(* CODESYS project festo_cmmt_as_etc.library
   DefaultNamespace: KOSTAL.TC3.Device.Axis.FESTO.CMMT_AS.ETC
   DocFormat: reStructuredText
   Description: Library to handle the FESTO CMMT_AS axis controller via EtherCAT
   Author: A.Zajic
   Title: KOSTAL.TC3.Device.Axis.FESTO.CMMT_AS.ETC
   Version: 2019.0.0.0
   Company: KOSTAL GmbH & Co.KG
   Placeholder: KOSTAL.TC3.Device.Axis.FESTO.CMMT_AS.ETC

Project tree, tasks and I/O mapping:
  libraries: Festo_PtP_Base, 3.5.15.32 (Festo); Festo_PtP_CiA402, 3.5.15.32 (Festo); Festo_PtP_CiA402_ETC, 3.5.15.32 (Festo); Festo_PtP_CiA402_ETC_CMMT_AS, 3.5.15.32 (Festo); Festo_PtP_Virtual, 3.5.15.32 (Festo); KOSTAL.TC3.Components.Stringhandler, 2019.1.1.0 (KOSTAL GmbH & Co.KG); KOSTAL.TC3.Core.plcResponse, 2019.0.1.0 (KOSTAL GmbH & Co.KG); KOSTAL.TC3.Core.process, 2019.3.0.0 (KOSTAL GmbH & Co.KG); KOSTAL.TC3.Device.Axis.I_LinearAxis, 2019.0.0.0 (KOSTAL GmbH & Co.KG); Tc2_Standard, 3.3.3.0 (Beckhoff Automation GmbH); Tc2_System, 3.4.24.0 (Beckhoff Automation GmbH); Tc3_Module, 3.3.21.0 (Beckhoff Automation GmbH)
  DUT/
    data type E_HomingMethod
  Interface/
    interface I_LinearAxis_position: IlinearAxis_Direction, IlinearAxis_FaultDescripition, IlinearAxis_HomingMethod, IlinearAxis_HomingPosition, IlinearAxis_isOn, IlinearAxis_Jerk, IlinearAxis_JogMode, IlinearAxis_MoveTorque, IlinearAxis_moveVelocity, IlinearAxis_RelativePos, IlinearAxis_SpeedAct, IlinearAxis_TorqueAct
  POE/
    COMMANDS/
      function block FB_EnableAxis [ST]: _isLinked, Enable, status, _FBmain, Execute, FBmain, link
      function block FB_homing [ST]: _a_finish, _a_home, _a_homing, _a_checkAxisEnabled, _a_init, _stepFail, _deviceDefine, _isLinked, HomingMethod, Position, Release, status, _FBmain, Execute, FBmain, link
      function block FB_move_Jog [ST]: _a_finish, _a_home, _a_checkAxisEnabled, _a_init, _a_jog, _stepFail, _deviceDefine, _isLinked, JogMode, jogNegative, jogPositive, Release, status, _FBmain, Execute, FBmain, link
      function block FB_move_Position [ST]: _a_finish, _a_home, _a_checkAxisEnabled, _a_init, _a_moveTo, _absoluteMotion, _relativeMotion, _stepFail, _deviceDefine, _isLinked, Accel, Decel, Direction, Jerk, Position, relativePos, Release, status, Velocity, _FBmain, Execute, FBmain, link
      function block FB_move_Record [ST]: _a_finish, _a_home, _a_checkAxisEnabled, _a_init, _a_moveTo, _stepFail, _deviceDefine, _isLinked, recordNo, Release, status, _FBmain, Execute, FBmain, link
      function block FB_move_Torque [ST]: _a_finish, _a_home, _a_checkAxisEnabled, _a_init, _a_moveTorque, _stepFail, _deviceDefine, _isLinked, Release, status, Torque, TorqueRamp, Velocity, _FBmain, Execute, FBmain, link
      function block FB_move_Velocity [ST]: _a_finish, _a_home, _a_checkAxisEnabled, _a_init, _a_moveVelo, _stepFail, _deviceDefine, _isLinked, Accel, Decel, Jerk, Release, status, Velocity, _FBmain, Execute, FBmain, link
      function block FB_Reset [ST]: _isLinked, Reset, status, _FBmain, Execute, FBmain, link
      function block FB_stopAxis [ST]: _a_home, _a_stopAxis, _stepFail, _deviceDefine, _isLinked, status, _FBmain, Execute, FBmain, link
    function block FB_FESTO_CMMT_AS [ST]: IlinearAxis_acceleration, IlinearAxis_deceleration, IlinearAxis_Direction, IlinearAxis_Fault, IlinearAxis_FaultDescripition, IlinearAxis_Homing, IlinearAxis_HomingMethod, IlinearAxis_HomingPosition, IlinearAxis_isOn, IlinearAxis_Jerk, IlinearAxis_JogMode, IlinearAxis_JogNegative_X, IlinearAxis_JogPositive_X, IlinearAxis_MoveRecord, IlinearAxis_MoveToPosition, IlinearAxis_MoveTorque, IlinearAxis_moveVelocity, IlinearAxis_Off, IlinearAxis_On, IlinearAxis_PositionAct, IlinearAxis_RelativePos, IlinearAxis_Release, IlinearAxis_ResetFault, IlinearAxis_Speed, IlinearAxis_SpeedAct, IlinearAxis_State, IlinearAxis_TorqueAct, _toggleGet, _FBmain, FBmain
  Project Information/
    function F_GetCompany [ST]
    function F_GetTitle [ST]
    function F_GetVersion [ST]
  Version/
    global variables Global_Version
*)

// DUT/E_HomingMethod
{attribute 'qualified_only'}
{attribute 'strict'}
TYPE E_HomingMethod :
(
	negStopLimSwitchWithTrToRefSw	:=-27,//-27; negative stop/limit switch with travel to reference switch
	posStopLimSwitchWithTrToRefSw	:=-23,//-23; positive stop/limit switch with travel to reference switch
	positiveStop					:=-18,//-18; positive stop
	negativeStop					:=-17,//-17; negative stop
	posStopWithZeroPls 				:= -2,//-2; positive stop with zero pulse
	negStopWithZeroPls 				:= -1,//-1; negative stop with zero pulse
	
	deviceSetting					:=  0,//0; homing method and axis zero point parametrised in the device are used
	
	negHwSwitchWithZeroPls 			:=  1,//1; negative HW limit switch with zero pulse
	posHwSwitchWithZeroPls 			:=  2,//2; positive HW limit switch with zero pulse
	posRefSwitchWithZeroPls			:=	7,//7; positive reference switch with zero pulse
	negRefSwitchWithZeroPls			:= 11,//11; negative reference switch with zero pulse
	negHwLimSwitch					:= 17,//17; negative HW limit switch
	posHwLimSwitch					:= 18,//18; positive HW limit switch
	posRefSwitch					:= 23,//23; positive reference switch
	negRefSwitch					:= 27,//27; negative reference switch
	currPosWithNegZeroPls			:= 33,//33; current position with negative zero pulse
	currPosWithPosZeroPls			:= 34,//34; current position with positive zero pulse
	currentPosition					:= 37 //37; current position (default setting)
)DINT;
END_TYPE

// Version/Global_Version
{attribute 'TcGenerated'}
{attribute 'no-analysis'}
{attribute 'linkalways'}
// This function has been automatically generated from the project information.
VAR_GLOBAL CONSTANT
	{attribute 'const_non_replaced'}
	stLibVersion_KOSTAL_TC3_Device_Axis_FESTO_CMMT_AS_ETC : ST_LibVersion := (iMajor := 2019, iMinor := 0, iBuild := 0, iRevision := 0, nFlags := 0, sVersion := '2019.0.0.0');
END_VAR

// Interface/I_LinearAxis_position
INTERFACE I_LinearAxis_position EXTENDS KOSTAL_TC3_Device_Axis_Interface.I_LinearAxis_position

(*
 defines the positioning direction if "modulo" is activated
*)
PROPERTY IlinearAxis_Direction : Festo_PtP_Base.MC_DIRECTION
GET
END_GET
SET
END_SET
END_PROPERTY

PROPERTY IlinearAxis_FaultDescripition : string(255);
GET
END_GET
END_PROPERTY

(*
 sets the homing method to CiA402 specification (see. the dirver documentation)
*)
PROPERTY IlinearAxis_HomingMethod : E_HomingMethod
GET
END_GET
SET
END_SET
END_PROPERTY

(*
 Absolute position if reference switch was detected
*)
PROPERTY IlinearAxis_HomingPosition : REAL
GET
END_GET
SET
END_SET
END_PROPERTY

(*
 Returns TRUE, if the axis is powered (drive is enabled)
 *)
PROPERTY IlinearAxis_isOn : bool
GET
END_GET
END_PROPERTY

(*
 jerk (in user units)
*)
PROPERTY IlinearAxis_Jerk : REAL
GET
END_GET
SET
END_SET
END_PROPERTY

(*
 0(mcDefault)=velo1 and velo2; 1(mcOnlyVelocity1); 2(mcOnlyVelocity2)
*)
PROPERTY IlinearAxis_JogMode : Festo_PtP_Base.MC_JOG_MODE
GET
END_GET
SET
END_SET
END_PROPERTY

(*
 Starts a motion with continuous torque measured at the motor shaft.
 The specified velocity is not exceeded.
*)
METHOD IlinearAxis_MoveTorque
VAR_INPUT
	Torque		: REAL; //setpoint torque at the motor shaft (in Nm)
	TorqueRamp	: REAL; //torque ramp (in Nm/s)
END_VAR
END_METHOD

(*
 Starts a controlled motion with a defined velocity.
 NOTE:
 If one of the inputs "Accel", "Decel" or "Jerk" = 0 when the motion starts, 
 the dynamic value set in the motor controller is used for this motion parameter.
*)
METHOD IlinearAxis_moveVelocity : REFERENCE TO KOSTAL_TC3_Core_plcResponse.FB_PlcResponse
VAR_INPUT
END_VAR
END_METHOD

(*
 Sets, if the position is relative or absolut
 TRUE=position is relative/ FALSE=position is absolute
*)
PROPERTY IlinearAxis_RelativePos : bool
GET
END_GET
SET
END_SET
END_PROPERTY

PROPERTY IlinearAxis_SpeedAct : REAL
GET
END_GET
END_PROPERTY

PROPERTY IlinearAxis_TorqueAct : REAL
GET
END_GET
END_PROPERTY

END_INTERFACE

// POE/COMMANDS/FB_EnableAxis
FUNCTION_BLOCK FB_EnableAxis

VAR
	// general
	_CMMT_AS		: REFERENCE TO Festo_PtP_CiA402_ETC_CMMT_AS.AXIS_REF_CiA402_ETC_CMMT_AS;
									
	_status			: KOSTAL_TC3_Core_plcResponse.FB_PlcResponse;
	_concat			: KOSTAL_TC3_Components_Stringhandler.FB_CONCAT;
	
	_Execute		: BOOL;
	_THIS_Called	: BOOL;

	// controll FB(s)
	_enableDrive	: Festo_PtP_Base.MC_Power_Festo;
	_enable			: BOOL;	
END_VAR

METHOD PROTECTED _isLinked : BOOL
VAR_INPUT
END_VAR

_isLinked:= __ISVALIDREF(_CMMT_AS);
END_METHOD

PROPERTY PUBLIC Enable : bool
GET
Enable:=_enable;
END_GET
SET
_enable:=Enable;
END_SET
END_PROPERTY

(*
| Function
| ========
| status of command execution
*)
PROPERTY PUBLIC status : REFERENCE TO KOSTAL_TC3_Core_plcResponse.FB_PlcResponse
GET


status REF= _status;
END_GET
END_PROPERTY

METHOD PROTECTED _FBmain
VAR_INPUT
END_VAR

_THIS_Called:= TRUE;

IF NOT _isLinked() THEN

	_status.clear();
	_status.fail:= TRUE;
	_status.description:= 'Reference to CMMT_ST is not valid';

	RETURN;

END_IF

IF NOT _execute THEN
	_status.clear();
	_status.ready:= TRUE;
END_IF

_enableDrive(
	Axis:= _CMMT_AS, 
	Enable:= _enable AND NOT _CMMT_AS.AxisError);
	
IF _CMMT_AS.AxisError THEN
	
	_status.clear();
	_status.finish:=TRUE;
	_status.fail:= TRUE;
	_status.description:='Enable Axis/ fault detect - try to reset';
	
ELSIF _enableDrive.Error THEN
	_status.clear();
	_status.finish:= TRUE;
	_status.fail:= TRUE;
	
	_concat.new(4);
	_concat.addContent(1, 'enable axis/ ErrID:');
	_concat.addContent(2, WORD_TO_STRING(_enableDrive.ErrorID));
	_concat.addContent(3, '/ ');
	_concat.addContent(4,_enableDrive.ErrorString );
	_status.description:= _concat.getResult();
	_concat.clear();
	
ELSIF NOT _enable AND NOT _enableDrive.Status AND _CMMT_AS.AxisState=AXIS_STATE.Disabled THEN
	_status.clear();
	_status.finish:= TRUE;
	_status.pass:= TRUE;
	_status.description:='axis is DISABLED';
	
ELSIF _enable AND _enableDrive.Status AND _enableDrive.Valid THEN
	_status.clear();
	_status.finish:= TRUE;
	_status.pass:= TRUE;
	_status.description:='axis is ENABLED';
	
ELSIF NOT _enable THEN
	_status.clear();
	_status.busy:= TRUE;
	_status.description:='axis will be DISABLED';
	
ELSIF _enable THEN
	_status.clear();
	_status.busy:= TRUE;
	_status.description:='axis will be ENABLED';	
END_IF
END_METHOD

METHOD PUBLIC Execute : BOOL

IF NOT _THIS_Called THEN

	_Execute:= TRUE;

	_FBmain();
	
	Execute:= _status.finish AND _status.pass;
	
END_IF
END_METHOD

METHOD PUBLIC FBmain
VAR_INPUT
END_VAR

IF NOT _THIS_Called THEN

	_Execute:= FALSE;

	_FBmain();
	
END_IF

_THIS_Called:= FALSE;
END_METHOD

METHOD PUBLIC link 

VAR_INPUT
	CMMT_AS	:	reference to Festo_PtP_CiA402_ETC_CMMT_AS.AXIS_REF_CiA402_ETC_CMMT_AS;
END_VAR

_CMMT_AS REF= CMMT_AS;
END_METHOD

END_FUNCTION_BLOCK

// POE/COMMANDS/FB_homing
FUNCTION_BLOCK FB_homing

VAR
	// general
	_CMMT_AS		: REFERENCE TO Festo_PtP_CiA402_ETC_CMMT_AS.AXIS_REF_CiA402_ETC_CMMT_AS;
	
	_step			: KOSTAL_TC3_Core_process.FB_processStep;
	_status			: KOSTAL_TC3_Core_plcResponse.FB_PlcResponse;
	_concat			: KOSTAL_TC3_Components_Stringhandler.FB_CONCAT;
	
	_Execute		: BOOL;
	_THIS_Called	: BOOL;
	
	_stop			: BOOL;
	_release		: BOOL;
	
	// controll FB(s)
	_homing			: Festo_PtP_Base.MC_Home_Festo;
	_stopAxis		: Festo_PtP_Base.MC_Stop_Festo;	
	
	// motion parameters
	_position		: REAL;
	_homingMethod	: E_HomingMethod:=0; 	
END_VAR

METHOD PROTECTED _a_finish
VAR_INPUT
END_VAR

(* result is set in the previous step *);
END_METHOD

METHOD PROTECTED _a_home
VAR_INPUT
END_VAR

IF NOT _Execute THEN
	
	_status.clear();
	_status.ready:= TRUE;

ELSE	

	_status.clear();
	_status.busy:= TRUE;

	_step.INC();	

END_IF
END_METHOD

METHOD PROTECTED _a_homing 
VAR
	_noFault 	: BOOL;
END_VAR
_homing.Execute:=TRUE;

IF _homing.Error THEN
	
	_status.clear();
	_status.finish:= TRUE;
	_status.fail:= TRUE;
	
	_concat.new(4);
	_concat.addContent(1, 'move home/ ErrID:');
	_concat.addContent(2, WORD_TO_STRING(_homing.ErrorID));
	_concat.addContent(3, '/ ');
	_concat.addContent(4,_homing.ErrorString );
	_status.description:= _concat.getResult();
	_concat.clear();
	
	_step.INC();
	
ELSIF _CMMT_AS.AxisError THEN
	
	_status.clear();
	_status.busy:=TRUE;
	_status.fail:= TRUE;
	
	_concat.new(4);
	_concat.addContent(1, 'move home/ ErrID:');
	_concat.addContent(2, WORD_TO_STRING(_CMMT_AS.AxisErrorID));
	_concat.addContent(3, '/ ');
	_concat.addContent(4,_CMMT_AS.AxisErrorString );
	_status.description:= _concat.getResult();
	_concat.clear();

	_step.INC();
	
ELSIF _CMMT_AS.AxisState=AXIS_STATE.ErrorStop OR _CMMT_AS.AxisState=AXIS_STATE.Stopping THEN
	_status.clear();
	_status.finish:= TRUE;
	_status.fail:= TRUE;
	_status.description:= 'homing was stopped';
		
	_step.INC();
	
ELSIF NOT _CMMT_AS.Enabled THEN
	
	_status.clear();
	_status.finish:= TRUE;
	_status.fail:= TRUE;
	_status.description:= 'Axis not ON';	

	_step.INC();
	
ELSIF NOT _release THEN 
	
	_status.clear();
	_status.finish:= TRUE;
	_status.fail:= TRUE;
	_status.description:= 'Axis not released';	

	_step.INC();
		
ELSIF _homing.Done THEN
	
	_status.clear();
	_status.finish:= TRUE;
	_status.pass:= TRUE;
	_status.description:= 'homing successfully executed';
	_step.INC();
	
ELSE
	_status.clear();
	_status.busy:= TRUE;
	_status.description:= 'wait for homing completed';	
END_IF
END_METHOD

METHOD PROTECTED _a_checkAxisEnabled
VAR_INPUT
END_VAR
IF _CMMT_AS.Enabled THEN
	_step.INC();
	
ELSE
	_status.clear();
	_status.busy:= TRUE;
	_status.description:='wait for axis enabled';
END_IF
END_METHOD

METHOD PROTECTED _a_init
VAR_INPUT
END_VAR
IF _CMMT_AS.AxisError THEN
	
	_status.clear();
	_status.busy:=TRUE;
	_status.fail:= TRUE;
	
	_concat.new(4);
	_concat.addContent(1, 'fault detect - try to reset/ ErrID:');
	_concat.addContent(2, WORD_TO_STRING(_CMMT_AS.AxisErrorID));
	_concat.addContent(3, '/ ');
	_concat.addContent(4,_CMMT_AS.AxisErrorString );
	_status.description:= _concat.getResult();
	_concat.clear();

ELSIF NOT _CMMT_AS.Enabled THEN
	
	_status.clear();
	_status.busy:= TRUE;
	_status.description:= 'Waiting for axis ON (drive is not ON)';
	
ELSIF NOT _release THEN
	
	_status.clear();
	_status.busy:= TRUE;
	_status.description:= 'Wating for axis released';
	
ELSIF _CMMT_AS.IsMoving THEN
	
	_status.clear();
	_status.busy:= TRUE;
	_status.description:= 'Waiting for another moving completed';

ELSE
	_step.INC();
END_IF
END_METHOD

METHOD PROTECTED _stepFail
VAR_INPUT
END_VAR

_status.clear();
_status.fail:= TRUE;
_concat.new(3);
_concat.addContent(1, 'Step: ');
_concat.addContent(2, INT_TO_STRING(_step.actual));
_concat.addContent(3, ' does not exist');
_status.description:= _concat.getResult();
_concat.clear();
END_METHOD

METHOD PROTECTED _deviceDefine
VAR_INPUT
END_VAR
_homing(
	Axis:= _CMMT_AS, 
	Position:= _position, 
	HomingMethod:= _homingMethod );
_homing.Execute:=FALSE;

// stop the axis if the command is not called before finished
IF (NOT _Execute OR NOT _release) AND _homing.Active THEN
	_stop:=TRUE;
END_IF
_stopAxis(
	Axis:= _CMMT_AS, 
	Execute:= _stop, 
	Done=> , 
	Busy=> , 
	CommandAborted=> , 
	Error=> , 
	ErrorID=> , 
	ErrorString=> );
IF _stopAxis.Done THEN
	_stop:=FALSE;
END_IF
END_METHOD

METHOD PROTECTED _isLinked : BOOL
VAR_INPUT
END_VAR

_isLinked:= __ISVALIDREF(_CMMT_AS);
END_METHOD

PROPERTY PUBLIC HomingMethod : E_HomingMethod
GET
HomingMethod:=_homingMethod;
END_GET
SET
_homingMethod:=HomingMethod;
END_SET
END_PROPERTY

PROPERTY PUBLIC Position : real
GET
Position:=_position;
END_GET
SET
_position:=_Position;
END_SET
END_PROPERTY

PROPERTY PUBLIC Release : bool
GET
Release:=_release;
END_GET
SET
_release:=Release;
END_SET
END_PROPERTY

(*
| Function
| ========
| status of command execution
*)
PROPERTY PUBLIC status : REFERENCE TO KOSTAL_TC3_Core_plcResponse.FB_PlcResponse
GET


status REF= _status;
END_GET
END_PROPERTY

METHOD PROTECTED _FBmain
VAR_INPUT
END_VAR

_THIS_Called:= TRUE;

IF NOT _isLinked() THEN

	_status.clear();
	_status.fail:= TRUE;
	_status.description:= 'Reference to CMMT_ST is not valid';
	_step.init();

	RETURN;

END_IF


IF NOT _Execute  AND (_step.actual <> 0) THEN _step.init();END_IF

_step.Header();

CASE _step.actual OF

	0:	_a_home();
	
	1:	_a_init();
	2:	_a_checkAxisEnabled();
	3:	_a_homing();
	
	4:	_a_finish();
	
ELSE
	
	_stepFail();
		
END_CASE

_deviceDefine();
END_METHOD

METHOD PUBLIC Execute : BOOL

IF NOT _THIS_Called THEN

	_Execute:= TRUE;

	_FBmain();
	
	Execute:= _status.finish AND _status.pass;
	
END_IF
END_METHOD

METHOD PUBLIC FBmain
VAR_INPUT
END_VAR

IF NOT _THIS_Called THEN

	_Execute:= FALSE;

	_FBmain();
	
END_IF

_THIS_Called:= FALSE;
END_METHOD

METHOD PUBLIC link 

VAR_INPUT
	CMMT_AS	:	reference to Festo_PtP_CiA402_ETC_CMMT_AS.AXIS_REF_CiA402_ETC_CMMT_AS;
END_VAR

_CMMT_AS REF= CMMT_AS;
END_METHOD

END_FUNCTION_BLOCK

// POE/COMMANDS/FB_move_Jog
FUNCTION_BLOCK FB_move_Jog

VAR
	// general
	_CMMT_AS		: REFERENCE TO Festo_PtP_CiA402_ETC_CMMT_AS.AXIS_REF_CiA402_ETC_CMMT_AS;
	
	_step			: KOSTAL_TC3_Core_process.FB_processStep;
	_status			: KOSTAL_TC3_Core_plcResponse.FB_PlcResponse;
	_concat			: KOSTAL_TC3_Components_Stringhandler.FB_CONCAT;
	
	_Execute		: BOOL;
	_THIS_Called	: BOOL;
	
	_release		: BOOL;
	
	// controll FB(s)
	_moveJog		: Festo_PtP_Base.MC_Jog_Festo;
	
	// motion parametes
	_jogMode		: Festo_PtP_Base.MC_JOG_MODE:=MC_JOG_MODE.mcDefault;
	_jogPositive	: BOOL;
	_jogNegative	: BOOL;
END_VAR

METHOD PROTECTED _a_finish
VAR_INPUT
END_VAR

(* result is set in the previous step *);
END_METHOD

METHOD PROTECTED _a_home
VAR_INPUT
END_VAR

(*IF NOT  _CMMT_AS.HomingValid THEN

	_status.clear();
	_status.fail:= TRUE;
	_status.finish:=TRUE;
	_status.description:= 'NOT referenced, homing necessary';
		
ELS*)IF NOT _Execute THEN
	
	_status.clear();
	_status.ready:= TRUE;

ELSE	

	_status.clear();
	_status.busy:= TRUE;

	_step.INC();	

END_IF
END_METHOD

METHOD PROTECTED _a_checkAxisEnabled
VAR_INPUT
END_VAR
IF _CMMT_AS.Enabled THEN
	_step.INC();
	
ELSE
	_status.clear();
	_status.busy:= TRUE;
	_status.description:='wait for axis enabled';
END_IF
END_METHOD

METHOD PROTECTED _a_init
VAR_INPUT
END_VAR
IF _CMMT_AS.AxisError THEN
	
	_status.clear();
	_status.busy:=TRUE;
	_status.fail:= TRUE;
	
	_concat.new(4);
	_concat.addContent(1, 'fault detect - try to reset/ ErrID:');
	_concat.addContent(2, WORD_TO_STRING(_CMMT_AS.AxisErrorID));
	_concat.addContent(3, '/ ');
	_concat.addContent(4,_CMMT_AS.AxisErrorString );
	_status.description:= _concat.getResult();
	_concat.clear();
	
ELSIF NOT _CMMT_AS.Enabled THEN
	
	_status.clear();
	_status.busy:= TRUE;
	_status.description:= 'Waiting for axis ON (drive is not ON)';
	
ELSIF NOT _release THEN
	
	_status.clear();
	_status.busy:= TRUE;
	_status.description:= 'Wating for axis released';
	
ELSIF _CMMT_AS.IsMoving THEN
	
	_status.clear();
	_status.busy:= TRUE;
	_status.description:= 'Waiting for another moving completed';

ELSE
	_step.INC();
END_IF
END_METHOD

METHOD PROTECTED _a_jog 
VAR
	_noFault 	: BOOL;
END_VAR
_moveJog.JogNegative:=_jogNegative AND NOT _jogPositive;
_moveJog.JogPositive:=_jogPositive AND NOT _jogNegative;


IF _moveJog.Error THEN
	
	_status.clear();
	_status.finish:= TRUE;
	_status.fail:= TRUE;
	
	_concat.new(4);
	_concat.addContent(1, 'move JOG/ ErrID:');
	_concat.addContent(2, WORD_TO_STRING(_moveJog.ErrorID));
	_concat.addContent(3, '/ ');
	_concat.addContent(4,_moveJog.ErrorString );
	_status.description:= _concat.getResult();
	_concat.clear();
	
	_step.INC();

ELSIF _CMMT_AS.AxisError THEN
	
	_status.clear();
	_status.busy:=TRUE;
	_status.fail:= TRUE;
	
	_concat.new(4);
	_concat.addContent(1, 'move JOG/ ErrID:');
	_concat.addContent(2, WORD_TO_STRING(_CMMT_AS.AxisErrorID));
	_concat.addContent(3, '/ ');
	_concat.addContent(4,_CMMT_AS.AxisErrorString );
	_status.description:= _concat.getResult();
	_concat.clear();

	_step.INC();
	
ELSIF NOT _CMMT_AS.Enabled THEN
	
	_status.clear();
	_status.finish:= TRUE;
	_status.fail:= TRUE;
	_status.description:= 'Axis not ON';	

	_step.INC();	
ELSIF NOT _release THEN 
	
	_status.clear();
	_status.finish:= TRUE;
	_status.fail:= TRUE;
	_status.description:= 'Axis not released';	

	_step.INC();	
	
ELSE
	_status.clear();
	_status.busy:= TRUE;
	IF _jogNegative THEN
		_status.description:= 'Axis: JOG-';
	ELSIF _jogPositive THEN
		_status.description:= 'Axis: JOG+';
	ELSE
		_status.description:= 'Axis: no JOG is active';
	END_IF
END_IF
END_METHOD

METHOD PROTECTED _stepFail
VAR_INPUT
END_VAR

_status.clear();
_status.fail:= TRUE;
_concat.new(3);
_concat.addContent(1, 'Step: ');
_concat.addContent(2, INT_TO_STRING(_step.actual));
_concat.addContent(3, ' does not exist');
_status.description:= _concat.getResult();
_concat.clear();
END_METHOD

METHOD PROTECTED _deviceDefine
VAR_INPUT
END_VAR
_moveJog(	Axis:= _CMMT_AS, 
			JogMode:= _jogMode, 
			ErrorID=> , 
			ErrorString=> );
_moveJog.JogNegative:=FALSE;
_moveJog.JogPositive:=FALSE;
END_METHOD

METHOD PROTECTED _isLinked : BOOL
VAR_INPUT
END_VAR

_isLinked:= __ISVALIDREF(_CMMT_AS);
END_METHOD

PROPERTY PUBLIC JogMode :  Festo_PtP_Base.MC_JOG_MODE
GET
JogMode :=_jogMode;
END_GET
SET
_jogMode:=JogMode;
END_SET
END_PROPERTY

(*
| As long as the value is TRUE, the selected axis is moving in negative direction
*)
PROPERTY PUBLIC jogNegative : BOOL
GET

jogNegative:= _jogNegative;
END_GET
SET

_jogNegative:= jogNegative;
END_SET
END_PROPERTY

(*
| As long as the value is TRUE, the selected axis is moving in positive direction
*)
PROPERTY PUBLIC jogPositive : BOOL
GET

jogPositive:= _jogPositive;
END_GET
SET

_jogPositive:= jogPositive;
END_SET
END_PROPERTY

PROPERTY PUBLIC Release : bool
GET
Release:=_release;
END_GET
SET
_release:=Release;
END_SET
END_PROPERTY

(*
| Function
| ========
| status of command execution
*)
PROPERTY PUBLIC status : REFERENCE TO KOSTAL_TC3_Core_plcResponse.FB_PlcResponse
GET


status REF= _status;
END_GET
END_PROPERTY

METHOD PROTECTED _FBmain
VAR_INPUT
END_VAR

_THIS_Called:= TRUE;

IF NOT _isLinked() THEN

	_status.clear();
	_status.fail:= TRUE;
	_status.description:= 'Reference to CMMT_ST is not valid';
	_step.init();

	RETURN;

END_IF


IF NOT _Execute  AND (_step.actual <> 0) THEN _step.init();END_IF

_step.Header();

CASE _step.actual OF

	0:	_a_home();
	
	1:	_a_init();
	2:	_a_checkAxisEnabled();
	3:	_a_jog();
	
	4:	_a_finish();
	
ELSE
	
	_stepFail();
		
END_CASE

_deviceDefine();
END_METHOD

METHOD PUBLIC Execute : BOOL

IF NOT _THIS_Called THEN

	_Execute:= TRUE;

	_FBmain();
	
	Execute:= _status.finish AND _status.pass;
	
END_IF
END_METHOD

METHOD PUBLIC FBmain
VAR_INPUT
END_VAR

IF NOT _THIS_Called THEN

	_Execute:= FALSE;

	_FBmain();
	
END_IF

_THIS_Called:= FALSE;
END_METHOD

METHOD PUBLIC link 

VAR_INPUT
	CMMT_AS	:	reference to Festo_PtP_CiA402_ETC_CMMT_AS.AXIS_REF_CiA402_ETC_CMMT_AS;
END_VAR

_CMMT_AS REF= CMMT_AS;
END_METHOD

END_FUNCTION_BLOCK

// POE/COMMANDS/FB_move_Position
FUNCTION_BLOCK FB_move_Position

VAR
	// general
	_CMMT_AS		: REFERENCE TO Festo_PtP_CiA402_ETC_CMMT_AS.AXIS_REF_CiA402_ETC_CMMT_AS;
	
	_step			: KOSTAL_TC3_Core_process.FB_processStep;
	_status			: KOSTAL_TC3_Core_plcResponse.FB_PlcResponse;
	_concat			: KOSTAL_TC3_Components_Stringhandler.FB_CONCAT;
	
	_Execute		: BOOL;
	_THIS_Called	: BOOL;
	
	_release		: BOOL;
	_stop			: BOOL;
	
	// controll FB(s)	
	_moveAbs		: Festo_PtP_Base.MC_MoveAbsolute_Festo;
	_moveRel		: Festo_PtP_Base.MC_MoveRelative_Festo;
	_stopAxis		: Festo_PtP_Base.MC_Stop_Festo;	
	
	// motion parametes
	_relativePos	: BOOL;	// =FALSE : move absolute position/ =TRUE : relative position
	_position		: REAL;	// position in user unit
	_velocity		: REAL;	// velocity 
	_accel			: REAL; // acceleration
	_decel			: REAL; // deceleration
	_jerk			: REAL;
	_direction		: Festo_PtP_Base.MC_DIRECTION:=MC_DIRECTION.mcNormal;
END_VAR

METHOD PROTECTED _a_finish
VAR_INPUT
END_VAR

(* result is set in the previous step *);
END_METHOD

METHOD PROTECTED _a_home
VAR_INPUT
END_VAR
IF NOT  _CMMT_AS.HomingValid THEN

	_status.clear();
	_status.fail:= TRUE;
	_status.finish:=TRUE;
	_status.description:= 'NOT referenced, homing necessary';
	
ELSIF NOT _Execute THEN
	
	_status.clear();
	_status.ready:= TRUE;

ELSE	

	_status.clear();
	_status.busy:= TRUE;

	_step.INC();	

END_IF
END_METHOD

METHOD PROTECTED _a_checkAxisEnabled
VAR_INPUT
END_VAR
IF _CMMT_AS.Enabled THEN
	_step.INC();
	
ELSE
	_status.clear();
	_status.busy:= TRUE;
	_status.description:='wait for axis enabled';
END_IF
END_METHOD

METHOD PROTECTED _a_init
VAR_INPUT
END_VAR
IF _CMMT_AS.AxisError THEN
	
	_status.clear();
	_status.busy:=TRUE;
	_status.fail:= TRUE;
	
	_concat.new(4);
	_concat.addContent(1, 'fault detect - try to reset/ ErrID:');
	_concat.addContent(2, WORD_TO_STRING(_CMMT_AS.AxisErrorID));
	_concat.addContent(3, '/ ');
	_concat.addContent(4,_CMMT_AS.AxisErrorString );
	_status.description:= _concat.getResult();
	_concat.clear();
	
ELSIF NOT _CMMT_AS.Enabled THEN
	
	_status.clear();
	_status.busy:= TRUE;
	_status.description:= 'Waiting for axis ON (drive is not ON)';
	
ELSIF NOT _release THEN
	
	_status.clear();
	_status.busy:= TRUE;
	_status.description:= 'Wating for axis released';
	
ELSIF _CMMT_AS.IsMoving THEN
	
	_status.clear();
	_status.busy:= TRUE;
	_status.description:= 'Waiting for another moving completed';

ELSE
	_step.INC();
END_IF
END_METHOD

METHOD PROTECTED _a_moveTo 
VAR
	_noFault 	: BOOL;
END_VAR
IF _relativePos THEN
	_relativeMotion();
ELSE
	_absoluteMotion();
END_IF
END_METHOD

METHOD PROTECTED _absoluteMotion 
VAR
	_noFault 	: BOOL;
END_VAR
_moveAbs.Execute:=TRUE;

IF _moveAbs.Error THEN
	
	_status.clear();
	_status.finish:= TRUE;
	_status.fail:= TRUE;
	
	_concat.new(4);
	_concat.addContent(1, 'move absolut/ ErrID:');
	_concat.addContent(2, WORD_TO_STRING(_moveAbs.ErrorID));
	_concat.addContent(3, '/ ');
	_concat.addContent(4,_moveAbs.ErrorString );
	_status.description:= _concat.getResult();
	_concat.clear();
	
	_step.INC();

ELSIF _CMMT_AS.AxisError THEN
	
	_status.clear();
	_status.busy:=TRUE;
	_status.fail:= TRUE;
	
	_concat.new(4);
	_concat.addContent(1, 'move absolut/ ErrID:');
	_concat.addContent(2, WORD_TO_STRING(_CMMT_AS.AxisErrorID));
	_concat.addContent(3, '/ ');
	_concat.addContent(4,_CMMT_AS.AxisErrorString );
	_status.description:= _concat.getResult();
	_concat.clear();

	_step.INC();
	
ELSIF _CMMT_AS.AxisState=AXIS_STATE.ErrorStop OR _CMMT_AS.AxisState=AXIS_STATE.Stopping THEN
	_status.clear();
	_status.finish:= TRUE;
	_status.fail:= TRUE;
	_status.description:= 'moving was stopped before target reached';
		
	_step.INC();

ELSIF NOT _CMMT_AS.Enabled THEN
	
	_status.clear();
	_status.finish:= TRUE;
	_status.fail:= TRUE;
	_status.description:= 'Axis not ON';	

	_step.INC();
	
ELSIF NOT _release THEN 
	
	_status.clear();
	_status.finish:= TRUE;
	_status.fail:= TRUE;
	_status.description:= 'Axis not released';	

	_step.INC();
			
ELSIF _moveAbs.Done THEN
	_status.clear();
	_status.pass:= TRUE;
	_status.finish:= TRUE;
	_status.description:= 'motion is completed';
	_step.INC();

ELSE	
	_status.clear();
	_status.busy:= TRUE;
	_status.description:= 'wait for motion completed';	
END_IF
END_METHOD

METHOD PROTECTED _relativeMotion 
VAR
	_noFault 	: BOOL;
END_VAR
_moveRel.Execute:=TRUE;

IF _moveRel.Error THEN
	
	_status.clear();
	_status.finish:= TRUE;
	_status.fail:= TRUE;
	
	_concat.new(4);
	_concat.addContent(1, 'move relative/ ErrID:');
	_concat.addContent(2, WORD_TO_STRING(_moveRel.ErrorID));
	_concat.addContent(3, '/ ');
	_concat.addContent(4,_moveRel.ErrorString );
	_status.description:= _concat.getResult();
	_concat.clear();
	
	_step.INC();

ELSIF _CMMT_AS.AxisError THEN
	
	_status.clear();
	_status.busy:=TRUE;
	_status.fail:= TRUE;
	
	_concat.new(4);
	_concat.addContent(1, 'move relative/ ErrID:');
	_concat.addContent(2, WORD_TO_STRING(_CMMT_AS.AxisErrorID));
	_concat.addContent(3, '/ ');
	_concat.addContent(4,_CMMT_AS.AxisErrorString );
	_status.description:= _concat.getResult();
	_concat.clear();

	_step.INC();
	
ELSIF _CMMT_AS.AxisState=AXIS_STATE.ErrorStop OR _CMMT_AS.AxisState=AXIS_STATE.Stopping THEN
	_status.clear();
	_status.finish:= TRUE;
	_status.fail:= TRUE;
	_status.description:= 'moving was stopped before target reached';
		
	_step.INC();

ELSIF NOT _CMMT_AS.Enabled THEN
	
	_status.clear();
	_status.finish:= TRUE;
	_status.fail:= TRUE;
	_status.description:= 'Axis not ON';	

	_step.INC();
	
ELSIF NOT _release THEN 
	
	_status.clear();
	_status.finish:= TRUE;
	_status.fail:= TRUE;
	_status.description:= 'Axis not released';	

	_step.INC();
				
ELSIF _moveRel.Done THEN
	_status.clear();
	_status.pass:= TRUE;
	_status.finish:= TRUE;
	_status.description:= 'motion is completed';
	_step.INC();

ELSE	
	_status.clear();
	_status.busy:= TRUE;
	_status.description:= 'wait for motion completed';	
END_IF
END_METHOD

METHOD PROTECTED _stepFail
VAR_INPUT
END_VAR

_status.clear();
_status.fail:= TRUE;
_concat.new(3);
_concat.addContent(1, 'Step: ');
_concat.addContent(2, INT_TO_STRING(_step.actual));
_concat.addContent(3, ' does not exist');
_status.description:= _concat.getResult();
_concat.clear();
END_METHOD

METHOD PROTECTED _deviceDefine
VAR_INPUT
END_VAR
_moveAbs(	Axis:= _CMMT_AS,  
			Position:= _position, 
			Velocity:= _velocity, 
			Acceleration:= _accel, 
			Deceleration:= _decel, 
			Jerk:= _jerk, 
			Direction:= _direction, 
			BufferMode:= MC_BUFFER_MODE.mcAborting );
_moveAbs.Execute:=FALSE;

_moveRel(
	Axis:= _CMMT_AS, 
	Distance:= _position, 
	Velocity:= _velocity, 
	Acceleration:= _accel, 
	Deceleration:= _decel, 
	Jerk:= _jerk, 
	Direction:= _direction, 
	BufferMode:= MC_BUFFER_MODE.mcAborting );
_moveRel.Execute:=FALSE;

// stop the axis if the command is not called before finished
IF (NOT _Execute OR NOT _release) AND (_moveAbs.Active OR _moveRel.Active) THEN
	_stop:=TRUE;
END_IF
_stopAxis(
	Axis:= _CMMT_AS, 
	Execute:= _stop, 
	Done=> , 
	Busy=> , 
	CommandAborted=> , 
	Error=> , 
	ErrorID=> , 
	ErrorString=> );
IF _stopAxis.Done THEN
	_stop:=FALSE;
END_IF
END_METHOD

METHOD PROTECTED _isLinked : BOOL
VAR_INPUT
END_VAR

_isLinked:= __ISVALIDREF(_CMMT_AS);
END_METHOD

PROPERTY PUBLIC Accel : real
GET
Accel:=_accel;
END_GET
SET
_accel:=Accel;
END_SET
END_PROPERTY

PROPERTY PUBLIC Decel : real
GET
Decel:=_decel;
END_GET
SET
_decel:=Decel;
END_SET
END_PROPERTY

PROPERTY PUBLIC Direction : Festo_PtP_Base.MC_DIRECTION
GET
Direction:=_direction;
END_GET
SET
_direction:=Direction;
END_SET
END_PROPERTY

PROPERTY PUBLIC Jerk : real
GET
Jerk:=_jerk;
END_GET
SET
_jerk:=Jerk;
END_SET
END_PROPERTY

PROPERTY PUBLIC Position : real
GET
Position:=_position;
END_GET
SET
_position:=Position;
END_SET
END_PROPERTY

(*
| Function
| ========
| Definition if the position is relative/absolute
| TRUE = position will be relative to the last setpoint value
| FALSE = position will be absolute
*)
PROPERTY PUBLIC relativePos : bool
GET
relativePos:=_relativePos;
END_GET
SET
_relativePos:=relativePos;
END_SET
END_PROPERTY

PROPERTY PUBLIC Release : bool
GET
Release:=_release;
END_GET
SET
_release:=Release;
END_SET
END_PROPERTY

(*
| Function
| ========
| status of command execution
*)
PROPERTY PUBLIC status : REFERENCE TO KOSTAL_TC3_Core_plcResponse.FB_PlcResponse
GET


status REF= _status;
END_GET
END_PROPERTY

PROPERTY PUBLIC Velocity : real
GET
Velocity:=_velocity;
END_GET
SET
_velocity:=Velocity;
END_SET
END_PROPERTY

METHOD PROTECTED _FBmain
VAR_INPUT
END_VAR

_THIS_Called:= TRUE;

IF NOT _isLinked() THEN

	_status.clear();
	_status.fail:= TRUE;
	_status.description:= 'Reference to CMMT_ST is not valid';
	_step.init();

	RETURN;

END_IF

_CMMT_AS();

IF NOT _Execute  AND (_step.actual <> 0) THEN _step.init();END_IF

_step.Header();

CASE _step.actual OF

	0:	_a_home();
	
	1:	_a_init();
	2:	_a_checkAxisEnabled();
	3:	_a_moveTo();

	4:	_a_finish();
	
ELSE
	
	_stepFail();
		
END_CASE

_deviceDefine();
END_METHOD

METHOD PUBLIC Execute : BOOL

IF NOT _THIS_Called THEN

	_Execute:= TRUE;

	_FBmain();
	
	Execute:= _status.finish AND _status.pass;
	
END_IF
END_METHOD

METHOD PUBLIC FBmain
VAR_INPUT
END_VAR

IF NOT _THIS_Called THEN

	_Execute:= FALSE;

	_FBmain();
	
END_IF

_THIS_Called:= FALSE;
END_METHOD

METHOD PUBLIC link 

VAR_INPUT
	CMMT_AS	:	reference to Festo_PtP_CiA402_ETC_CMMT_AS.AXIS_REF_CiA402_ETC_CMMT_AS;
END_VAR

_CMMT_AS REF= CMMT_AS;
END_METHOD

END_FUNCTION_BLOCK

// POE/COMMANDS/FB_move_Record
FUNCTION_BLOCK FB_move_Record

VAR
	// general
	_CMMT_AS		: REFERENCE TO Festo_PtP_CiA402_ETC_CMMT_AS.AXIS_REF_CiA402_ETC_CMMT_AS;
	
	_step			: KOSTAL_TC3_Core_process.FB_processStep;
	_status			: KOSTAL_TC3_Core_plcResponse.FB_PlcResponse;
	_concat			: KOSTAL_TC3_Components_Stringhandler.FB_CONCAT;
	
	_Execute		: BOOL;
	_THIS_Called	: BOOL;
	
	_stop			: BOOL;
	_release		: BOOL;
	
	// controll FB(s)
	_moveRecord		: Festo_PtP_Base.MC_RecordTable_Festo;
	_stopAxis		: Festo_PtP_Base.MC_Stop_Festo;	
	
	// motion parametes
	_recordNo		: DINT;
END_VAR

METHOD PROTECTED _a_finish
VAR_INPUT
END_VAR

(* result is set in the previous step *);
END_METHOD

METHOD PROTECTED _a_home
VAR_INPUT
END_VAR

IF NOT  _CMMT_AS.HomingValid THEN

	_status.clear();
	_status.fail:= TRUE;
	_status.finish:=TRUE;
	_status.description:= 'NOT referenced, homing necessary';
	
ELSIF NOT _Execute THEN
	
	_status.clear();
	_status.ready:= TRUE;

ELSE	

	_status.clear();
	_status.busy:= TRUE;

	_step.INC();	

END_IF
END_METHOD

METHOD PROTECTED _a_checkAxisEnabled
VAR_INPUT
END_VAR
IF _CMMT_AS.Enabled THEN
	_step.INC();
	
ELSE
	_status.clear();
	_status.busy:= TRUE;
	_status.description:='wait for axis enabled';
END_IF
END_METHOD

METHOD PROTECTED _a_init
VAR_INPUT
END_VAR
IF _CMMT_AS.AxisError THEN
	
	_status.clear();
	_status.busy:=TRUE;
	_status.fail:= TRUE;
	
	_concat.new(4);
	_concat.addContent(1, 'fault detect - try to reset/ ErrID:');
	_concat.addContent(2, WORD_TO_STRING(_CMMT_AS.AxisErrorID));
	_concat.addContent(3, '/ ');
	_concat.addContent(4,_CMMT_AS.AxisErrorString );
	_status.description:= _concat.getResult();
	_concat.clear();
	
ELSIF NOT _CMMT_AS.Enabled THEN
	
	_status.clear();
	_status.busy:= TRUE;
	_status.description:= 'Waiting for axis ON (drive is not ON)';
	
ELSIF NOT _release THEN
	
	_status.clear();
	_status.busy:= TRUE;
	_status.description:= 'Wating for axis released';
	
ELSIF _CMMT_AS.IsMoving THEN
	
	_status.clear();
	_status.busy:= TRUE;
	_status.description:= 'Waiting for another moving completed';

ELSE
	_step.INC();
END_IF
END_METHOD

METHOD PROTECTED _a_moveTo 
VAR
	_noFault 	: BOOL;
END_VAR
_moveRecord.Execute:=TRUE;

IF _moveRecord.Error<>0 THEN
	
	_status.clear();
	_status.finish:= TRUE;
	_status.fail:= TRUE;
	
	_concat.new(4);
	_concat.addContent(1, 'move record/ ErrID:');
	_concat.addContent(2, WORD_TO_STRING(_moveRecord.ErrorID));
	_concat.addContent(3, '/ ');
	_concat.addContent(4,_moveRecord.ErrorString );
	_status.description:= _concat.getResult();
	_concat.clear();
	
	_step.INC();

ELSIF _CMMT_AS.AxisError THEN
	
	_status.clear();
	_status.busy:=TRUE;
	_status.fail:= TRUE;
	
	_concat.new(4);
	_concat.addContent(1, 'move record/ ErrID:');
	_concat.addContent(2, WORD_TO_STRING(_CMMT_AS.AxisErrorID));
	_concat.addContent(3, '/ ');
	_concat.addContent(4,_CMMT_AS.AxisErrorString );
	_status.description:= _concat.getResult();
	_concat.clear();

	_step.INC();

ELSIF _CMMT_AS.AxisState=AXIS_STATE.ErrorStop OR _CMMT_AS.AxisState=AXIS_STATE.Stopping THEN
	_status.clear();
	_status.finish:= TRUE;
	_status.fail:= TRUE;
	_status.description:= 'moving was stopped before target reached';
		
	_step.INC();

	ELSIF NOT _CMMT_AS.Enabled THEN
	
	_status.clear();
	_status.finish:= TRUE;
	_status.fail:= TRUE;
	_status.description:= 'Axis not ON';	

	_step.INC();
	
ELSIF NOT _release THEN 
	
	_status.clear();
	_status.finish:= TRUE;
	_status.fail:= TRUE;
	_status.description:= 'Axis not released';	

	_step.INC();
				
ELSIF _moveRecord.Done THEN
	
	_status.clear();
	_status.pass:= TRUE;
	_status.finish:= TRUE;
	_status.description:= 'motion is completed';
	_step.INC();
	
ELSE
	_status.clear();
	_status.busy:= TRUE;
	_status.description:= 'wait for moving completed';	
END_IF
END_METHOD

METHOD PROTECTED _stepFail
VAR_INPUT
END_VAR

_status.clear();
_status.fail:= TRUE;
_concat.new(3);
_concat.addContent(1, 'Step: ');
_concat.addContent(2, INT_TO_STRING(_step.actual));
_concat.addContent(3, ' does not exist');
_status.description:= _concat.getResult();
_concat.clear();
END_METHOD

METHOD PROTECTED _deviceDefine
VAR_INPUT
END_VAR
_moveRecord(
	Axis:= _CMMT_AS, 
	RecordNumber:= _recordNo, 
	BufferMode:= MC_BUFFER_MODE.mcAborting);
_moveRecord.Execute:=FALSE;

// stop the axis if the command is not called before finished
IF (NOT _Execute OR NOT _release) AND _moveRecord.Active THEN
	_stop:=TRUE;
END_IF
_stopAxis(
	Axis:= _CMMT_AS, 
	Execute:= _stop, 
	Done=> , 
	Busy=> , 
	CommandAborted=> , 
	Error=> , 
	ErrorID=> , 
	ErrorString=> );
IF _stopAxis.Done THEN
	_stop:=FALSE;
END_IF
END_METHOD

METHOD PROTECTED _isLinked : BOOL
VAR_INPUT
END_VAR

_isLinked:= __isvalidref(_CMMT_AS);
END_METHOD

(*
| Function
| ========
| Record number
*)
PROPERTY PUBLIC recordNo : DINT
GET

recordNo:= _recordNo;
END_GET
SET

_recordNo:= recordNo;
END_SET
END_PROPERTY

PROPERTY PUBLIC Release : bool
GET
Release:=_release;
END_GET
SET
_release:=Release;
END_SET
END_PROPERTY

(*
| Function
| ========
| status of command execution
*)
PROPERTY PUBLIC status : REFERENCE TO KOSTAL_TC3_Core_plcResponse.FB_PlcResponse
GET


status REF= _status;
END_GET
END_PROPERTY

METHOD PROTECTED _FBmain
VAR_INPUT
END_VAR

_THIS_Called:= TRUE;

IF NOT _isLinked() THEN

	_status.clear();
	_status.fail:= TRUE;
	_status.description:= 'Reference to CMMT_ST is not valid';
	_step.init();

	RETURN;

END_IF


IF NOT _Execute  AND (_step.actual <> 0) THEN _step.init();END_IF

_step.Header();

CASE _step.actual OF

	0:	_a_home();
	
	1:	_a_init();
	2:	_a_checkAxisEnabled();
	3:	_a_moveTo();
	
	4:	_a_finish();
	
ELSE
	
	_stepFail();
		
END_CASE

_deviceDefine();
END_METHOD

METHOD PUBLIC Execute : BOOL

IF NOT _THIS_Called THEN

	_Execute:= TRUE;

	_FBmain();
	
	Execute:= _status.finish AND _status.pass;
	
END_IF
END_METHOD

METHOD PUBLIC FBmain
VAR_INPUT
END_VAR

IF NOT _THIS_Called THEN

	_Execute:= FALSE;

	_FBmain();
	
END_IF

_THIS_Called:= FALSE;
END_METHOD

METHOD PUBLIC link 

VAR_INPUT
	CMMT_AS	:	reference to Festo_PtP_CiA402_ETC_CMMT_AS.AXIS_REF_CiA402_ETC_CMMT_AS;
END_VAR

_CMMT_AS REF= CMMT_AS;
END_METHOD

END_FUNCTION_BLOCK

// POE/COMMANDS/FB_move_Torque
FUNCTION_BLOCK FB_move_Torque

VAR
	// general
	_CMMT_AS		: REFERENCE TO Festo_PtP_CiA402_ETC_CMMT_AS.AXIS_REF_CiA402_ETC_CMMT_AS;
	
	_step			: KOSTAL_TC3_Core_process.FB_processStep;
	_status			: KOSTAL_TC3_Core_plcResponse.FB_PlcResponse;
	_concat			: KOSTAL_TC3_Components_Stringhandler.FB_CONCAT;
	
	_Execute		: BOOL;
	_THIS_Called	: BOOL;
	
	_stop			: BOOL;
	_release		: BOOL;
	
	// controll FB(s)
	_moveTorque		: Festo_PtP_Base.MC_TorqueControl_Festo;
	_stopAxis		: Festo_PtP_Base.MC_Stop_Festo;	

	
	// motion parametes
	_velocity		: REAL;	// velocity 
	_torque			: REAL;
	_torqueRamp		: REAL;
END_VAR

METHOD PROTECTED _a_finish
VAR_INPUT
END_VAR

(* result is set in the previous step *);
END_METHOD

METHOD PROTECTED _a_home
VAR_INPUT
END_VAR

IF NOT  _CMMT_AS.HomingValid THEN

	_status.clear();
	_status.fail:= TRUE;
	_status.finish:=TRUE;
	_status.description:= 'NOT referenced, homing necessary';
	
ELSIF NOT _Execute THEN
	
	_status.clear();
	_status.ready:= TRUE;

ELSE	

	_status.clear();
	_status.busy:= TRUE;

	_step.INC();	

END_IF
END_METHOD

METHOD PROTECTED _a_checkAxisEnabled
VAR_INPUT
END_VAR
IF _CMMT_AS.Enabled THEN
	_step.INC();
	
ELSE
	_status.clear();
	_status.busy:= TRUE;
	_status.description:='wait for axis enabled';
END_IF
END_METHOD

METHOD PROTECTED _a_init
VAR_INPUT
END_VAR
IF _CMMT_AS.AxisError THEN
	
	_status.clear();
	_status.busy:=TRUE;
	_status.fail:= TRUE;
	
	_concat.new(4);
	_concat.addContent(1, 'fault detect - try to reset/ ErrID:');
	_concat.addContent(2, WORD_TO_STRING(_CMMT_AS.AxisErrorID));
	_concat.addContent(3, '/ ');
	_concat.addContent(4,_CMMT_AS.AxisErrorString );
	_status.description:= _concat.getResult();
	_concat.clear();
	
ELSIF NOT _CMMT_AS.Enabled THEN
	
	_status.clear();
	_status.busy:= TRUE;
	_status.description:= 'Waiting for axis ON (drive is not ON)';
	
ELSIF NOT _release THEN
	
	_status.clear();
	_status.busy:= TRUE;
	_status.description:= 'Wating for axis released';
	
ELSIF _CMMT_AS.IsMoving THEN
	
	_status.clear();
	_status.busy:= TRUE;
	_status.description:= 'Waiting for another moving completed';

ELSE
	_step.INC();
END_IF
END_METHOD

METHOD PROTECTED _a_moveTorque 
VAR
	_noFault 	: BOOL;
END_VAR
_moveTorque.Execute:=TRUE;

IF _moveTorque.Error THEN
	
	_status.clear();
	_status.finish:= TRUE;
	_status.fail:= TRUE;
	
	_concat.new(4);
	_concat.addContent(1, 'move torque/ ErrID:');
	_concat.addContent(2, WORD_TO_STRING(_moveTorque.ErrorID));
	_concat.addContent(3, '/ ');
	_concat.addContent(4,_moveTorque.ErrorString );
	_status.description:= _concat.getResult();
	_concat.clear();
	
	_step.INC();

ELSIF _CMMT_AS.AxisError THEN
	
	_status.clear();
	_status.busy:=TRUE;
	_status.fail:= TRUE;
	
	_concat.new(4);
	_concat.addContent(1, 'move torque/ ErrID:');
	_concat.addContent(2, WORD_TO_STRING(_CMMT_AS.AxisErrorID));
	_concat.addContent(3, '/ ');
	_concat.addContent(4,_CMMT_AS.AxisErrorString );
	_status.description:= _concat.getResult();
	_concat.clear();

	_step.INC();
	
ELSIF _CMMT_AS.AxisState=AXIS_STATE.ErrorStop OR _CMMT_AS.AxisState=AXIS_STATE.Stopping THEN
	_status.clear();
	_status.finish:= TRUE;
	_status.fail:= TRUE;
	_status.description:= 'moving was stopped before target reached';
		
	_step.INC();

ELSIF NOT _CMMT_AS.Enabled THEN
	
	_status.clear();
	_status.finish:= TRUE;
	_status.fail:= TRUE;
	_status.description:= 'Axis not ON';	

	_step.INC();
	
ELSIF NOT _release THEN 
	
	_status.clear();
	_status.finish:= TRUE;
	_status.fail:= TRUE;
	_status.description:= 'Axis not released';	

	_step.INC();
				
ELSIF _moveTorque.InTorque THEN

	_status.clear();
	_status.pass:= TRUE;
	_status.finish:= TRUE;
	_status.description:= 'torque reached';
	_step.INC();

ELSE
	_status.clear();
	_status.busy:= TRUE;
	_status.description:= 'moving to requested torque ...';	
END_IF
END_METHOD

METHOD PROTECTED _stepFail
VAR_INPUT
END_VAR

_status.clear();
_status.fail:= TRUE;
_concat.new(3);
_concat.addContent(1, 'Step: ');
_concat.addContent(2, INT_TO_STRING(_step.actual));
_concat.addContent(3, ' does not exist');
_status.description:= _concat.getResult();
_concat.clear();
END_METHOD

METHOD PROTECTED _deviceDefine
VAR_INPUT
END_VAR
_moveTorque(
	Axis:= _CMMT_AS, 
	Torque:= _torque, 
	TorqueRamp:= _torqueRamp, 
	Velocity:= _velocity, 
	BufferMode:= MC_BUFFER_MODE.mcAborting );
_moveTorque.Execute:=FALSE;	

// stop the axis if the command is not called before finished
IF (NOT _Execute OR NOT _release) AND _moveTorque.Active THEN
	_stop:=TRUE;
END_IF
_stopAxis(
	Axis:= _CMMT_AS, 
	Execute:= _stop, 
	Done=> , 
	Busy=> , 
	CommandAborted=> , 
	Error=> , 
	ErrorID=> , 
	ErrorString=> );
IF _stopAxis.Done THEN
	_stop:=FALSE;
END_IF
END_METHOD

METHOD PROTECTED _isLinked : BOOL
VAR_INPUT
END_VAR

_isLinked:= __isvalidref(_CMMT_AS);
END_METHOD

PROPERTY PUBLIC Release : bool
GET
Release:=_release;
END_GET
SET
_release:=Release;
END_SET
END_PROPERTY

(*
| Function
| ========
| status of command execution
*)
PROPERTY PUBLIC status : REFERENCE TO KOSTAL_TC3_Core_plcResponse.FB_PlcResponse
GET


status REF= _status;
END_GET
END_PROPERTY

PROPERTY PUBLIC Torque : real
GET
Torque:=_torque;
END_GET
SET
_torque:=Torque;
END_SET
END_PROPERTY

PROPERTY PUBLIC TorqueRamp : real
GET
TorqueRamp:=_torqueRamp;
END_GET
SET
_torqueRamp:=TorqueRamp;
END_SET
END_PROPERTY

PROPERTY PUBLIC Velocity : real
GET
Velocity:=_velocity;
END_GET
SET
_velocity:=Velocity;
END_SET
END_PROPERTY

METHOD PROTECTED _FBmain
VAR_INPUT
END_VAR

_THIS_Called:= TRUE;

IF NOT _isLinked() THEN

	_status.clear();
	_status.fail:= TRUE;
	_status.description:= 'Reference to CMMT_ST is not valid';
	_step.init();

	RETURN;

END_IF


IF NOT _Execute  AND (_step.actual <> 0) THEN _step.init();END_IF

_step.Header();

CASE _step.actual OF

	0:	_a_home();
	
	1:	_a_init();
	2:	_a_checkAxisEnabled();
	3:	_a_moveTorque();
	
	4:	_a_finish();
	
ELSE
	
	_stepFail();
		
END_CASE

_deviceDefine();
END_METHOD

METHOD PUBLIC Execute : BOOL

IF NOT _THIS_Called THEN

	_Execute:= TRUE;

	_FBmain();
	
	Execute:= _status.finish AND _status.pass;
	
END_IF
END_METHOD

METHOD PUBLIC FBmain
VAR_INPUT
END_VAR

IF NOT _THIS_Called THEN

	_Execute:= FALSE;

	_FBmain();
	
END_IF

_THIS_Called:= FALSE;
END_METHOD

METHOD PUBLIC link 

VAR_INPUT
	CMMT_AS	:	reference to Festo_PtP_CiA402_ETC_CMMT_AS.AXIS_REF_CiA402_ETC_CMMT_AS;
END_VAR

_CMMT_AS REF= CMMT_AS;
END_METHOD

END_FUNCTION_BLOCK

// POE/COMMANDS/FB_move_Velocity
FUNCTION_BLOCK FB_move_Velocity

VAR
	// general
	_CMMT_AS		: REFERENCE TO Festo_PtP_CiA402_ETC_CMMT_AS.AXIS_REF_CiA402_ETC_CMMT_AS;
	
	_step			: KOSTAL_TC3_Core_process.FB_processStep;
	_status			: KOSTAL_TC3_Core_plcResponse.FB_PlcResponse;
	_concat			: KOSTAL_TC3_Components_Stringhandler.FB_CONCAT;
	
	_Execute		: BOOL;
	_THIS_Called	: BOOL;
	
	_stop			: BOOL;
	_release		: BOOL;

	// controll FB(s)
	_moveVelocity	: Festo_PtP_Base.MC_MoveVelocity_Festo;
	_stopAxis		: Festo_PtP_Base.MC_Stop_Festo;	

	// motion parametes
	_velocity		: REAL;	// velocity 
	_accel			: REAL; // acceleration
	_decel			: REAL; // deceleration
	_jerk			: REAL;
END_VAR

METHOD PROTECTED _a_finish
VAR_INPUT
END_VAR

(* result is set in the previous step *);
END_METHOD

METHOD PROTECTED _a_home
VAR_INPUT
END_VAR

IF NOT  _CMMT_AS.HomingValid THEN

	_status.clear();
	_status.fail:= TRUE;
	_status.finish:=TRUE;
	_status.description:= 'NOT referenced, homing necessary';
	
ELSIF NOT _Execute THEN
	
	_status.clear();
	_status.ready:= TRUE;

ELSE	

	_status.clear();
	_status.busy:= TRUE;

	_step.INC();	

END_IF
END_METHOD

METHOD PROTECTED _a_checkAxisEnabled
VAR_INPUT
END_VAR
IF _CMMT_AS.Enabled THEN
	_step.INC();
	
ELSE
	_status.clear();
	_status.busy:= TRUE;
	_status.description:='wait for axis enabled';
END_IF
END_METHOD

METHOD PROTECTED _a_init
VAR_INPUT
END_VAR
IF _CMMT_AS.AxisError THEN
	
	_status.clear();
	_status.busy:=TRUE;
	_status.fail:= TRUE;
	
	_concat.new(4);
	_concat.addContent(1, 'fault detect - try to reset/ ErrID:');
	_concat.addContent(2, WORD_TO_STRING(_CMMT_AS.AxisErrorID));
	_concat.addContent(3, '/ ');
	_concat.addContent(4,_CMMT_AS.AxisErrorString );
	_status.description:= _concat.getResult();
	_concat.clear();
	
ELSIF NOT _CMMT_AS.Enabled THEN
	
	_status.clear();
	_status.busy:= TRUE;
	_status.description:= 'Waiting for axis ON (drive is not ON)';
	
ELSIF NOT _release THEN
	
	_status.clear();
	_status.busy:= TRUE;
	_status.description:= 'Wating for axis released';
	
ELSIF _CMMT_AS.IsMoving THEN
	
	_status.clear();
	_status.busy:= TRUE;
	_status.description:= 'Waiting for another moving completed';

ELSE
	_step.INC();
END_IF
END_METHOD

METHOD PROTECTED _a_moveVelo 
VAR
	_noFault 	: BOOL;
END_VAR
_moveVelocity.Execute:=TRUE;

IF _moveVelocity.Error THEN
	
	_status.clear();
	_status.finish:= TRUE;
	_status.fail:= TRUE;
	
	_concat.new(4);
	_concat.addContent(1, 'move velocity/ ErrID:');
	_concat.addContent(2, WORD_TO_STRING(_moveVelocity.ErrorID));
	_concat.addContent(3, '/ ');
	_concat.addContent(4,_moveVelocity.ErrorString );
	_status.description:= _concat.getResult();
	_concat.clear();
	
	_step.INC();

ELSIF _CMMT_AS.AxisError THEN
	
	_status.clear();
	_status.busy:=TRUE;
	_status.fail:= TRUE;
	
	_concat.new(4);
	_concat.addContent(1, 'move velocity/ ErrID:');
	_concat.addContent(2, WORD_TO_STRING(_CMMT_AS.AxisErrorID));
	_concat.addContent(3, '/ ');
	_concat.addContent(4,_CMMT_AS.AxisErrorString );
	_status.description:= _concat.getResult();
	_concat.clear();

	_step.INC();

ELSIF _CMMT_AS.AxisState=AXIS_STATE.ErrorStop OR _CMMT_AS.AxisState=AXIS_STATE.Stopping THEN
	_status.clear();
	_status.finish:= TRUE;
	_status.fail:= TRUE;
	_status.description:= 'moving was stopped before target reached';
		
	_step.INC();

ELSIF NOT _CMMT_AS.Enabled THEN
	
	_status.clear();
	_status.finish:= TRUE;
	_status.fail:= TRUE;
	_status.description:= 'Axis not ON';	

	_step.INC();
	
ELSIF NOT _release THEN 
	
	_status.clear();
	_status.finish:= TRUE;
	_status.fail:= TRUE;
	_status.description:= 'Axis not released';	

	_step.INC();
				
ELSIF _moveVelocity.InVelocity THEN

	_status.clear();
	_status.pass:= TRUE;
	_status.finish:= TRUE;
	_status.description:= 'velocity reached';
	_step.INC();

ELSE
	_status.clear();
	_status.busy:= TRUE;
	_status.description:= 'moving to requested velocity ...';	
END_IF
END_METHOD

METHOD PROTECTED _stepFail
VAR_INPUT
END_VAR

_status.clear();
_status.fail:= TRUE;
_concat.new(3);
_concat.addContent(1, 'Step: ');
_concat.addContent(2, INT_TO_STRING(_step.actual));
_concat.addContent(3, ' does not exist');
_status.description:= _concat.getResult();
_concat.clear();
END_METHOD

METHOD PROTECTED _deviceDefine
VAR_INPUT
END_VAR
_moveVelocity(
	Axis:= _CMMT_AS, 
	Velocity:= _velocity, 
	Acceleration:= _accel, 
	Deceleration:= _decel, 
	Jerk:= _jerk, 
	BufferMode:=  MC_BUFFER_MODE.mcAborting );
_moveVelocity.Execute:=FALSE;

// stop the axis if the command is not called before finished
IF (NOT _Execute OR NOT _release) AND _moveVelocity.Active  THEN
	_stop:=TRUE;
END_IF
_stopAxis(
	Axis:= _CMMT_AS, 
	Execute:= _stop, 
	Done=> , 
	Busy=> , 
	CommandAborted=> , 
	Error=> , 
	ErrorID=> , 
	ErrorString=> );
IF _stopAxis.Done THEN
	_stop:=FALSE;
END_IF
END_METHOD

METHOD PROTECTED _isLinked : BOOL
VAR_INPUT
END_VAR

_isLinked:= __isvalidref(_CMMT_AS);
END_METHOD

PROPERTY PUBLIC Accel : real
GET
Accel:=_accel;
END_GET
SET
_accel:=Accel;
END_SET
END_PROPERTY

PROPERTY PUBLIC Decel : real
GET
Decel:=_decel;
END_GET
SET
_decel:=Decel;
END_SET
END_PROPERTY

PROPERTY PUBLIC Jerk : real
GET
Jerk:=_jerk;
END_GET
SET
_jerk:=Jerk;
END_SET
END_PROPERTY

PROPERTY PUBLIC Release : bool
GET
Release:=_release;
END_GET
SET
_release:=Release;
END_SET
END_PROPERTY

(*
| Function
| ========
| status of command execution
*)
PROPERTY PUBLIC status : REFERENCE TO KOSTAL_TC3_Core_plcResponse.FB_PlcResponse
GET


status REF= _status;
END_GET
END_PROPERTY

PROPERTY PUBLIC Velocity : real
GET
Velocity:=_velocity;
END_GET
SET
_velocity:=Velocity;
END_SET
END_PROPERTY

METHOD PROTECTED _FBmain
VAR_INPUT
END_VAR

_THIS_Called:= TRUE;

IF NOT _isLinked() THEN

	_status.clear();
	_status.fail:= TRUE;
	_status.description:= 'Reference to CMMT_ST is not valid';
	_step.init();

	RETURN;

END_IF


IF NOT _Execute  AND (_step.actual <> 0) THEN _step.init();END_IF

_step.Header();

CASE _step.actual OF

	0:	_a_home();
	
	1:	_a_init();
	2:	_a_checkAxisEnabled();
	3:	_a_moveVelo();
	
	4:	_a_finish();
	
ELSE
	
	_stepFail();
		
END_CASE

_deviceDefine();
END_METHOD

METHOD PUBLIC Execute : BOOL

IF NOT _THIS_Called THEN

	_Execute:= TRUE;

	_FBmain();
	
	Execute:= _status.finish AND _status.pass;
	
END_IF
END_METHOD

METHOD PUBLIC FBmain
VAR_INPUT
END_VAR

IF NOT _THIS_Called THEN

	_Execute:= FALSE;

	_FBmain();
	
END_IF

_THIS_Called:= FALSE;
END_METHOD

METHOD PUBLIC link 

VAR_INPUT
	CMMT_AS	:	reference to Festo_PtP_CiA402_ETC_CMMT_AS.AXIS_REF_CiA402_ETC_CMMT_AS;
END_VAR

_CMMT_AS REF= CMMT_AS;
END_METHOD

END_FUNCTION_BLOCK

// POE/COMMANDS/FB_Reset
FUNCTION_BLOCK FB_Reset

VAR
	// general
	_CMMT_AS		: REFERENCE TO Festo_PtP_CiA402_ETC_CMMT_AS.AXIS_REF_CiA402_ETC_CMMT_AS;
	
	_status			: KOSTAL_TC3_Core_plcResponse.FB_PlcResponse;
	_concat			: KOSTAL_TC3_Components_Stringhandler.FB_CONCAT;
	
	_Execute		: BOOL;
	_THIS_Called	: BOOL;

	// controll FB(s)
	_resetDrive		: Festo_PtP_Base.MC_Reset_Festo;
	_reset			: BOOL;	
END_VAR

METHOD PROTECTED _isLinked : BOOL
VAR_INPUT
END_VAR

_isLinked:= __ISVALIDREF(_CMMT_AS);
END_METHOD

PROPERTY PUBLIC Reset : bool
GET
Reset:=_reset;
END_GET
SET
_reset:=Reset;
END_SET
END_PROPERTY

(*
| Function
| ========
| status of command execution
*)
PROPERTY PUBLIC status : REFERENCE TO KOSTAL_TC3_Core_plcResponse.FB_PlcResponse
GET


status REF= _status;
END_GET
END_PROPERTY

METHOD PROTECTED _FBmain
VAR_INPUT
END_VAR

_THIS_Called:= TRUE;

IF NOT _isLinked() THEN

	_status.clear();
	_status.fail:= TRUE;
	_status.description:= 'Reference to CMMT_ST is not valid';

	RETURN;

END_IF

IF NOT _execute THEN
	_status.clear();
	_status.ready:= TRUE;
END_IF

_resetDrive(
	Axis:= _CMMT_AS, 
	Execute:= _reset, 
	Done=> , 
	Busy=> , 
	Error=> , 
	ErrorID=> , 
	ErrorString=> );
	
IF _resetDrive.Error THEN
	_status.clear();
	_status.finish:= TRUE;
	_status.fail:= TRUE;
	
	_concat.new(4);
	_concat.addContent(1, 'reset axis/ ErrID:');
	_concat.addContent(2, WORD_TO_STRING(_resetDrive.ErrorID));
	_concat.addContent(3, '/ ');
	_concat.addContent(4,_resetDrive.ErrorString );
	_status.description:= _concat.getResult();
	_concat.clear();
	
ELSIF _reset AND _resetDrive.Busy THEN
	_status.clear();
	_status.finish:= TRUE;
	_status.pass:= TRUE;
	_status.description:='axis error will be reseted';
	
ELSIF _reset AND _resetDrive.Done THEN
	_status.clear();
	_status.finish:= TRUE;
	_status.pass:= TRUE;
	_status.description:='reset axis error done';	
END_IF

_reset:=FALSE;
END_METHOD

METHOD PUBLIC Execute : BOOL

IF NOT _THIS_Called THEN

	_Execute:= TRUE;

	_FBmain();
	
	Execute:= _status.finish AND _status.pass;
	
END_IF
END_METHOD

METHOD PUBLIC FBmain
VAR_INPUT
END_VAR

IF NOT _THIS_Called THEN

	_Execute:= FALSE;

	_FBmain();
	
END_IF

_THIS_Called:= FALSE;
END_METHOD

METHOD PUBLIC link 

VAR_INPUT
	CMMT_AS	:	reference to Festo_PtP_CiA402_ETC_CMMT_AS.AXIS_REF_CiA402_ETC_CMMT_AS;
END_VAR

_CMMT_AS REF= CMMT_AS;
END_METHOD

END_FUNCTION_BLOCK

// POE/COMMANDS/FB_stopAxis
FUNCTION_BLOCK FB_stopAxis

VAR
	// general
	_CMMT_AS		: REFERENCE TO Festo_PtP_CiA402_ETC_CMMT_AS.AXIS_REF_CiA402_ETC_CMMT_AS;
	
	_step			: KOSTAL_TC3_Core_process.FB_processStep;
	_status			: KOSTAL_TC3_Core_plcResponse.FB_PlcResponse;
	_concat			: KOSTAL_TC3_Components_Stringhandler.FB_CONCAT;
	
	_Execute		: BOOL;
	_THIS_Called	: BOOL;

	// controll FB(s)
	_stopAxis	: Festo_PtP_Base.MC_Stop_Festo;	
END_VAR

METHOD PROTECTED _a_home
VAR_INPUT
END_VAR

IF NOT _Execute THEN
	
	_status.clear();
	_status.ready:= TRUE;

ELSE	

	_status.clear();
	_status.busy:= TRUE;

	_step.INC();	

END_IF
END_METHOD

METHOD PROTECTED _a_stopAxis
_stopAxis.Execute:=TRUE;

IF _stopAxis.Error<>0 THEN
	
	_status.clear();
	_status.fail:= TRUE;
	_status.finish:=TRUE;
	
	_concat.new(4);
	_concat.addContent(1, 'stop axis/ ErrID:');
	_concat.addContent(2, WORD_TO_STRING(_stopAxis.ErrorID));
	_concat.addContent(3, '/ ');
	_concat.addContent(4,_stopAxis.ErrorString );
	_status.description:= _concat.getResult();
	_concat.clear();

ELSIF NOT _stopAxis.Done THEN
	_status.clear();
	_status.pass:= TRUE;
	_status.finish:=TRUE;
	_status.description:='...stopped';
END_IF
END_METHOD

METHOD PROTECTED _stepFail
VAR_INPUT
END_VAR

_status.clear();
_status.fail:= TRUE;
_concat.new(3);
_concat.addContent(1, 'Step: ');
_concat.addContent(2, INT_TO_STRING(_step.actual));
_concat.addContent(3, ' does not exist');
_status.description:= _concat.getResult();
_concat.clear();
END_METHOD

METHOD PROTECTED _deviceDefine
VAR_INPUT
END_VAR
_stopAxis(Axis:= _CMMT_AS);
_stopAxis.Execute:=FALSE;
END_METHOD

METHOD PROTECTED _isLinked : BOOL
VAR_INPUT
END_VAR

_isLinked:= __ISVALIDREF(_CMMT_AS);
END_METHOD

(*
| Function
| ========
| status of command execution
*)
PROPERTY PUBLIC status : REFERENCE TO KOSTAL_TC3_Core_plcResponse.FB_PlcResponse
GET


status REF= _status;
END_GET
END_PROPERTY

METHOD PROTECTED _FBmain
VAR_INPUT
END_VAR

_THIS_Called:= TRUE;

IF NOT _isLinked() THEN

	_status.clear();
	_status.fail:= TRUE;
	_status.description:= 'Reference to CMMT_ST is not valid';
	_step.init();

	RETURN;

END_IF


IF NOT _Execute AND (_step.actual <> 0) THEN _step.init();	END_IF

_step.Header();

CASE _step.actual OF

	0:	_a_Home();
	
	1:	_a_stopAxis();
		
ELSE
	
	_stepFail();
		
END_CASE

_deviceDefine();
END_METHOD

METHOD PUBLIC Execute : BOOL

IF NOT _THIS_Called THEN

	_Execute:= TRUE;

	_FBmain();
	
	Execute:= _status.finish AND _status.pass;
	
END_IF
END_METHOD

METHOD PUBLIC FBmain
VAR_INPUT
END_VAR

IF NOT _THIS_Called THEN

	_Execute:= FALSE;

	_FBmain();
	
END_IF

_THIS_Called:= FALSE;
END_METHOD

METHOD PUBLIC link 

VAR_INPUT
	CMMT_AS	:	reference to Festo_PtP_CiA402_ETC_CMMT_AS.AXIS_REF_CiA402_ETC_CMMT_AS;
END_VAR

_CMMT_AS REF= CMMT_AS;
END_METHOD

END_FUNCTION_BLOCK

// POE/FB_FESTO_CMMT_AS
(*

:Author: Ales Zajic <a.zajic@kostal.com>
:Date: 2020-12-09

Function
==========
| Function block to control the axis controller FESTO CMMT-AS via EtherCAT
| It is a wrapper to the third party libraries (created by company FESTO)

IMPORTANT
=========
| The following third party libraries must be installed:
| Festo_PtP_Base
| Festo_PtP_CiA402
| Festo_PtP_CiA402_ETC
| Festo_PtP_CiA_ETC_CMMT_AS
| Festo_PtP_Virtual
| The third party libraries were created by company FESTO and they are free of charge available on their web-sides.
| Developed with the Festo-libraries version 3.5.15.32

Usage sample:
=============

.. code:: 

*)
FUNCTION_BLOCK FB_FESTO_CMMT_AS IMPLEMENTS I_LinearAxis_position,KOSTAL_TC3_Device_Axis_Interface.I_LinearAxis_jog,KOSTAL_TC3_Device_Axis_Interface.I_LinearAxis_record
VAR
	_CMMT_AS		: Festo_PtP_CiA402_ETC_CMMT_AS.AXIS_REF_CiA402_ETC_CMMT_AS;	
				
	_state			: KOSTAL_TC3_Core_plcResponse.FB_PlcResponse;
	_concat			: KOSTAL_TC3_Components_Stringhandler.FB_CONCAT;
	
	_enableAxis		: FB_EnableAxis;
	_stopAxis		: FB_stopAxis;
	_resetAxis		: FB_Reset;
	_homing			: FB_homing;
	_moveJog		: FB_move_Jog;
	_movePos		: FB_move_Position;
	_moveRecord		: FB_move_Record;
	_moveTorque		: FB_move_Torque;
	_moveVelocity	: FB_move_Velocity;	
	
	_toggle			: BOOL;
	_toggleTimer	: TON;
		
	_release		: BOOL;
	_isOn			: BOOL;
	
	_homingMethod	: E_HomingMethod:=E_HomingMethod.deviceSetting;//Homing method to CiA402 specification (see. the dirver documentation)
	_homing_Position: REAL;//Absolute position if reference switch was detected
	
	_jogMode		: Festo_PtP_Base.MC_JOG_MODE:=MC_JOG_MODE.mcDefault;// 0(mcDefault)=velo1 and velo2; 1(mcOnlyVelocity1); 2(mcOnlyVelocity2)
	
	_speed			: REAL;//maximum velocity (in user units)
	_accel			: REAL;//acceleration (in user units)
	_decel			: REAL;//deceleration (in user units)
	_jerk			: REAL;//jerk (in user units)
	_direction		: Festo_PtP_Base.MC_DIRECTION:=MC_DIRECTION.mcNormal;//defines the positioning direction if "modulo" is activated
	_relativePos	: BOOL;//TRUE the target position will be relative to the last set point/ FALSE the target position is absolute
END_VAR

(*
 sets the requested acceleration 
*)
PROPERTY IlinearAxis_acceleration : REAL
GET
IlinearAxis_acceleration:=_accel;
END_GET
SET
_accel:=IlinearAxis_acceleration;
END_SET
END_PROPERTY

(*
 sets the requested deceleration 
*)
PROPERTY IlinearAxis_deceleration : REAL
GET
IlinearAxis_deceleration:=_decel;
END_GET
SET
_decel:=IlinearAxis_deceleration;
END_SET
END_PROPERTY

(*
 defines the positioning direction if "modulo" is activated
*)
PROPERTY IlinearAxis_Direction : Festo_PtP_Base.MC_DIRECTION
GET
IlinearAxis_Direction:=_direction;
END_GET
SET
_direction:=IlinearAxis_Direction;
END_SET
END_PROPERTY

(*
 Returns TRUE, if the axis is in error
 *)
PROPERTY IlinearAxis_Fault : BOOL
GET
IlinearAxis_Fault:=_CMMT_AS.AxisError;
END_GET
END_PROPERTY

(*
| Returns the axis error ID and error description
*)
PROPERTY IlinearAxis_FaultDescripition : string(255);
GET
IF _CMMT_AS.AxisError THEN
	
	_concat.new(4);
	_concat.addContent(1, 'ErrID:');
	_concat.addContent(2, WORD_TO_STRING(_CMMT_AS.AxisErrorID));
	_concat.addContent(3, '/ ');
	_concat.addContent(4,_CMMT_AS.AxisErrorString );
	IlinearAxis_FaultDescripition :=_concat.getResult();
	_concat.clear();
	
ELSE
	IlinearAxis_FaultDescripition:='';
END_IF;
END_GET
END_PROPERTY

(*
 Executes referencing of the axis
 NOTE:
 If the "HomingMethod" input = 0, the homing method and axis zero point parameterised in the device are used. 
 The axis zero point specified in the block ("Position" input) is ignored. 
 If the "HomingMethod" input <> 0, the homing method and axis zero point parameterised in the device are overwritten.
*)
METHOD IlinearAxis_Homing : BOOL
_homing.HomingMethod:=_homingMethod;
_homing.Position:=_homing_Position;
_homing.Execute();

_state:=_homing.status;
IlinearAxis_Homing:=_homing.status.finish and _homing.status.pass;
END_METHOD

(*
 sets the homing method to CiA402 specification (see. the dirver documentation)
*)
PROPERTY IlinearAxis_HomingMethod : E_HomingMethod
GET
IlinearAxis_HomingMethod:=_homingMethod;
END_GET
SET
_homingMethod:=IlinearAxis_HomingMethod;
END_SET
END_PROPERTY

(*
 Absolute position if reference switch was detected
*)
PROPERTY IlinearAxis_HomingPosition : REAL
GET
IlinearAxis_HomingPosition:=_homing_Position;
END_GET
SET
_homing_Position:=IlinearAxis_HomingPosition;
END_SET
END_PROPERTY

(*
 Returns TRUE, if the axis is powered (drive is enabled)
 *)
PROPERTY IlinearAxis_isOn : bool
GET
IlinearAxis_isOn:=_isOn;
END_GET
END_PROPERTY

(*
 jerk (in user units)
*)
PROPERTY IlinearAxis_Jerk : REAL
GET
IlinearAxis_Jerk:=_jerk;
END_GET
SET
_jerk:=IlinearAxis_Jerk;
END_SET
END_PROPERTY

(*
 0(mcDefault)=velo1 and velo2; 1(mcOnlyVelocity1); 2(mcOnlyVelocity2)
*)
PROPERTY IlinearAxis_JogMode : Festo_PtP_Base.MC_JOG_MODE
GET
IlinearAxis_JogMode:=_jogMode;
END_GET
SET
_jogMode:=IlinearAxis_JogMode;
END_SET
END_PROPERTY

METHOD IlinearAxis_JogNegative_X
_moveJog.jogNegative:=TRUE;
_moveJog.jogPositive:=FALSE;
_moveJog.JogMode:=_jogMode;
_moveJog.Execute();

_state:=_moveJog.status;
END_METHOD

METHOD IlinearAxis_JogPositive_X
_moveJog.jogNegative:=FALSE;
_moveJog.jogPositive:=TRUE;
_moveJog.JogMode:=_jogMode;
_moveJog.Execute();

_state:=_moveJog.status;
END_METHOD

(*
 Executes the move defined in the selected record
*)
METHOD IlinearAxis_MoveRecord
VAR_INPUT
	recordNo	: UINT;
END_VAR
_moveRecord.recordNo:=recordNo;
_moveRecord.Execute();

_state:=_moveRecord.status;
END_METHOD

(*Move to given position*)
METHOD IlinearAxis_MoveToPosition
VAR_INPUT
	position	: REAL;
END_VAR
_movePos.Position:=position;
_movePos.Velocity:=_speed;
_movePos.Accel:=_accel;
_movePos.Decel:=_decel;
_movePos.Jerk:=_jerk;
_movePos.Direction:=_direction;
_movePos.relativePos:=_relativePos;
_movePos.Execute();

_state:=_movePos.status;
END_METHOD

(*
 Starts a motion with continuous torque measured at the motor shaft.
 The specified velocity is not exceeded.
*)
METHOD IlinearAxis_MoveTorque
VAR_INPUT
	Torque		: REAL; //setpoint torque at the motor shaft (in Nm)
	TorqueRamp	: REAL; //torque ramp (in Nm/s)
END_VAR
_moveTorque.Torque:=Torque;
_moveTorque.TorqueRamp:=TorqueRamp;
_moveTorque.Velocity:=_speed;
_moveTorque.Execute();

_state:=_moveTorque.status;
END_METHOD

(*
 Starts a controlled motion with a defined velocity.
 NOTE:
 If one of the inputs "Accel", "Decel" or "Jerk" = 0 when the motion starts, 
 the dynamic value set in the motor controller is used for this motion parameter.
*)
METHOD IlinearAxis_moveVelocity : REFERENCE TO KOSTAL_TC3_Core_plcResponse.FB_PlcResponse
VAR_INPUT
END_VAR
_moveVelocity.Velocity:=_speed;
_moveVelocity.Accel:=_accel;
_moveVelocity.Decel:=_decel;
_moveVelocity.Jerk:=_jerk;
_moveVelocity.Execute();

_state:=_moveVelocity.status;
END_METHOD

METHOD IlinearAxis_Off : BOOL
_enableAxis.Enable:=FALSE;
_enableAxis.Execute();

_state:=_enableAxis.status;
END_METHOD

METHOD IlinearAxis_On : BOOL
_enableAxis.Enable:=TRUE;
_enableAxis.Execute();

_state:=_enableAxis.status;
END_METHOD

PROPERTY IlinearAxis_PositionAct : REAL
GET
IlinearAxis_PositionAct:=_CMMT_AS.ActualPosition;
END_GET
END_PROPERTY

(*
 Sets, if the position is relative or absolut
 TRUE=position is relative/ FALSE=position is absolute
*)
PROPERTY IlinearAxis_RelativePos : bool
GET
IlinearAxis_RelativePos:=_relativePos;
END_GET
SET
_relativePos:=IlinearAxis_RelativePos;
END_SET
END_PROPERTY

METHOD IlinearAxis_Release : BOOL
VAR_INPUT
	release	: BOOL;
END_VAR
_release:=release;
END_METHOD

METHOD IlinearAxis_ResetFault : BOOL
_resetAxis.Reset:=_toggle;
_resetAxis.Execute();
END_METHOD

PROPERTY IlinearAxis_Speed : REAL
GET
IlinearAxis_Speed:=_speed;
END_GET
SET
_speed:=IlinearAxis_Speed;
END_SET
END_PROPERTY

PROPERTY IlinearAxis_SpeedAct : REAL
GET
IlinearAxis_SpeedAct:=_CMMT_AS.ActualVelocity;
END_GET
END_PROPERTY

PROPERTY IlinearAxis_State : REFERENCE TO KOSTAL_TC3_Device_Axis_Interface.KOSTAL_TC3_Core_plcResponse.FB_PlcResponse
GET
IlinearAxis_State ref=_state;
END_GET
END_PROPERTY

PROPERTY IlinearAxis_TorqueAct : REAL
GET
IlinearAxis_TorqueAct:=_CMMT_AS.ActualTorque;
END_GET
END_PROPERTY

METHOD PROTECTED _toggleGet
VAR_INPUT
END_VAR

IF NOT _toggleTimer.Q THEN
	_toggleTimer(IN:= TRUE, PT:= T#500MS);
ELSE
	_toggleTimer(IN:= FALSE);
	_toggle:= NOT _toggle;
END_IF
END_METHOD

METHOD PROTECTED _FBmain
VAR_INPUT
END_VAR
_state.clear();

_toggleGet();
_CMMT_AS();

_homing.link(_CMMT_AS);
_homing.Release:=_release;
_homing.FBmain();

_moveJog.link(_CMMT_AS);
_moveJog.FBmain();
_moveJog.Release:=_release;
_moveJog.jogNegative:=FALSE;
_moveJog.jogPositive:=FALSE;

_movePos.link(_CMMT_AS);
_movePos.Release:=_release;
_movePos.FBmain();

_moveRecord.link(_CMMT_AS);
_moveRecord.Release:=_release;
_moveRecord.FBmain();

_moveTorque.link(_CMMT_AS);
_moveTorque.Release:=_release;
_moveTorque.FBmain();

_moveVelocity.link(_CMMT_AS);
_moveVelocity.Release:=_release;	
_moveVelocity.FBmain();

_stopAxis.link(_CMMT_AS);
_stopAxis.FBmain();

_enableAxis.link(_CMMT_AS);
_enableAxis.FBmain();
_isOn:=_CMMT_AS.Enabled;

_resetAxis.link(_CMMT_AS);
_resetAxis.FBmain();
END_METHOD

METHOD PUBLIC FBmain
VAR_INPUT
END_VAR

_FBmain();
END_METHOD

END_FUNCTION_BLOCK

// Project Information/F_GetCompany
// This function has been automatically generated from the project information.
{attribute 'signature_flag' := '1073741824'}
{attribute 'TcGenerated'}
{attribute 'no-analysis'}
FUNCTION F_GetCompany : WSTRING
VAR_INPUT
	
END_VAR

F_GetCompany := "KOSTAL GmbH & Co.KG";

END_FUNCTION

// Project Information/F_GetTitle
// This function has been automatically generated from the project information.
{attribute 'signature_flag' := '1073741824'}
{attribute 'TcGenerated'}
{attribute 'no-analysis'}
FUNCTION F_GetTitle : WSTRING
VAR_INPUT
	
END_VAR

F_GetTitle := "KOSTAL.TC3.Device.Axis.FESTO.CMMT_AS.ETC";

END_FUNCTION

// Project Information/F_GetVersion
// This function has been automatically generated from the project information.
{attribute 'signature_flag' := '1073741824'}
{attribute 'TcGenerated'}
{attribute 'no-analysis'}
FUNCTION F_GetVersion : ST_LibVersion
VAR_INPUT
	
END_VAR

F_GetVersion.iMajor := 2019;
F_GetVersion.iMinor := 0;
F_GetVersion.iBuild := 0;
F_GetVersion.iRevision := 0;

END_FUNCTION
